FUNCTION_BLOCK MOD_OccupationLogic (* Decides Occupy and Release: occupy when free (or again by the owner), release only by the owner, and answer Accepted or an error code. Technical: Occupation by session ID: Occupy when free (or again by the owner), Release only by the owner *)
  (* Standard: 61499-2 *)
  (* Version 0.1, 2026-09-28, Project contributors, AAU Smart Production Lab *)
  PACKAGE modlib;
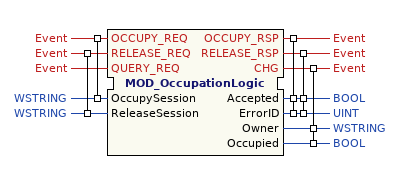
  EVENT_INPUT
    OCCUPY_REQ WITH OccupySession; (* Occupy(Session) was called *)
    RELEASE_REQ WITH ReleaseSession; (* Release(Session) was called *)
    QUERY_REQ; (* A block asks for the current owner *)
  END_EVENT
  EVENT_OUTPUT
    OCCUPY_RSP WITH Accepted, ErrorID; (* Answer to Occupy: Accepted, ErrorID *)
    RELEASE_RSP WITH Accepted, ErrorID; (* Answer to Release: Accepted, ErrorID *)
    CHG WITH Owner, Occupied; (* The value changed *)
  END_EVENT
  VAR_INPUT
    OccupySession : WSTRING; (* Session ID of the caller of Occupy *)
    ReleaseSession : WSTRING; (* Session ID of the caller of Release *)
  END_VAR
  VAR_OUTPUT
    Accepted : BOOL; (* The call was accepted *)
    ErrorID : UINT; (* Error code: 0 none, 1 PreconditionViolated, 2 InvariantViolated, 3 Timeout, 4 NotReady, 5 NotPermitted, 6 Busy, 7 Interrupted, 8 OutOfRange *)
    Owner : WSTRING; (* Session ID of the module's owner (empty: free) *)
    Occupied : BOOL; (* The module is occupied *)
  END_VAR
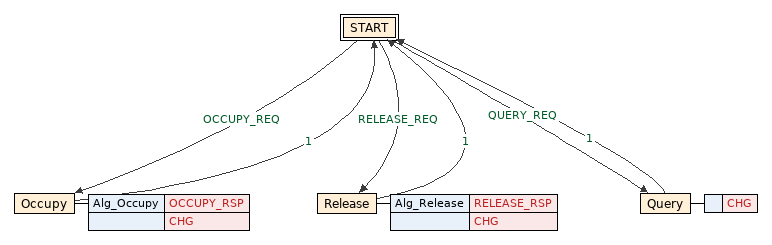
  EC_STATES
    START;
    Occupy : Alg_Occupy -> OCCUPY_RSP, -> CHG;
    Release : Alg_Release -> RELEASE_RSP, -> CHG;
    Query : -> CHG;
  END_STATES
  EC_TRANSITIONS
    START TO Occupy := OCCUPY_REQ;
    Occupy TO START := 1;
    START TO Release := RELEASE_REQ;
    Release TO START := 1;
    START TO Query := QUERY_REQ;
    Query TO START := 1;
  END_TRANSITIONS
  ALGORITHM Alg_Occupy IN ST:
IF (OccupySession <> "") AND ((Owner = "") OR (Owner = OccupySession)) THEN
  Owner := OccupySession;
  Occupied := TRUE;
  Accepted := TRUE;
  ErrorID := 0;
ELSE
  Accepted := FALSE;
  ErrorID := 5;
END_IF;
  END_ALGORITHM
  ALGORITHM Alg_Release IN ST:
IF (Owner <> "") AND (Owner = ReleaseSession) THEN
  Owner := "";
  Occupied := FALSE;
  Accepted := TRUE;
  ErrorID := 0;
ELSE
  Accepted := FALSE;
  ErrorID := 5;
END_IF;
  END_ALGORITHM
END_FUNCTION_BLOCK
